// TIA Portal V20 export
DATA_BLOCK "08_Systemzeit_DB"   // DB29
// stored: InstanceOfName 08_Systemzeit, InstanceOfType FB
"08_Systemzeit"
   // VAR
   //    outputTIME : Date_And_Time;
   //    returnValue : Int;
   //    inputTIME : Date_And_Time;
   //    returnValueT : Int;
   //    execute : Bool;
   // END_VAR
BEGIN
END_DATA_BLOCK
